(* Logix 5000 project; controller lab5BnB 5069-L306ERM rev 38.11; software revision 38.02 *)

TASK MainTask (periodic, rate 1 ms, priority 10, watchdog 1 ms) : MainProgram

MODULES
   Local : 5069-L306ERM (5069 0, rev 38.11)
       : 5069-OB16 (5069 2, rev 3.13, StandardDataDriven RPI 5 ms)
       : 5069-IB16 (5069 1, rev 2.16, StandardDataDriven RPI 5 ms)
       : vendor 1 type 115 code 320 (5069 4, rev 2.13, StandardDataDriven RPI 1 ms)
       : 5069-IF8 (5069 3, rev 3.11, StandardDataDriven RPI 1 ms)
END_MODULES

ADD_ON_INSTRUCTION Angle_Controller   (* revision 1.0 *)
VAR_INPUT
   Kp : REAL; {access None}
   Kd : REAL; {access None}
   Ki : REAL; {access None}
END_VAR
VAR_OUTPUT
   MotorInInt : REAL; {access None}
END_VAR
VAR_INPUT
   MotorVoltageInt : REAL; {access None}
   DesiredMotorAngleDeg : REAL; {access None}
END_VAR
VAR
   DERV_01 : DERIVATIVE := (Gain := 0.8, RTSTime := 1, DeltaT := 0.001);
   INTG_02 : INTEGRATOR := (IGain := 0.5, HighLimit := 4.0, LowLimit := -4.0, RTSTime := 1, Out := 1.9863874, DeltaT := 0.001);
   LPF_01 : FILTER_LOW_PASS := (WLag := 0.5, Order := 1, RTSTime := 1, DeltaT := 0.001);
   MUL_01 : FBD_MATH := (SourceA := 0.4);
   SCL_01 : SCALE := (In := 1.6115597, InRawMax := 2.8, InRawMin := -1.92, InEUMax := 90.0, InEUMin := -90.0, Limiting := 1, Out := 44.67813);
   SCL_02 : SCALE := (In := 1.9863874, InRawMax := 90.0, InRawMin := -90.0, InEUMax := -10.0, InEUMin := 10.0, Limiting := 1, Out := -0.2207098);
   SSUM_01 : SELECTED_SUMMER := (Gain1 := 1.0, Select1 := 1, Gain2 := 1.0, Select2 := 1, In3 := 1.9863874, Gain3 := 1.0, Select3 := 1, Gain4 := 1.0, Gain5 := 1.0, Gain6 := 1.0, Gain7 := 1.0, Gain8 := 1.0, Out := 1.9863874);
   SUB_01 : FBD_MATH := (SourceA := 45.0, SourceB := 45.0);
   BalanceMax : REAL := 2.8; {access None}
   BalanceMin : REAL := -1.92; {access None}
   MotorAngleDeg : REAL; {access None}
   MyError : REAL; {access None}
   PreFilter : REAL; {access None}
   PostFilter : REAL; {access None}
   __lECF02074BD2460E6 : REAL; {access None}
   __l28C6010D865A5A33 : REAL; {access None}
   __l0884565386038A91 : REAL; {access None}
   __l2DF07EE77D244EFB : REAL; {access None}
   __l1766871E0CB1B884 : REAL; {access None}
   __l0E750273472B5D8B : REAL; {access None}
   __lD887463BECBAFEBD : REAL; {access None}
   __l08A3F56F66BAD335 : REAL; {access None}
END_VAR

ROUTINE Logic   (* function block diagram *)
   SHEET 1
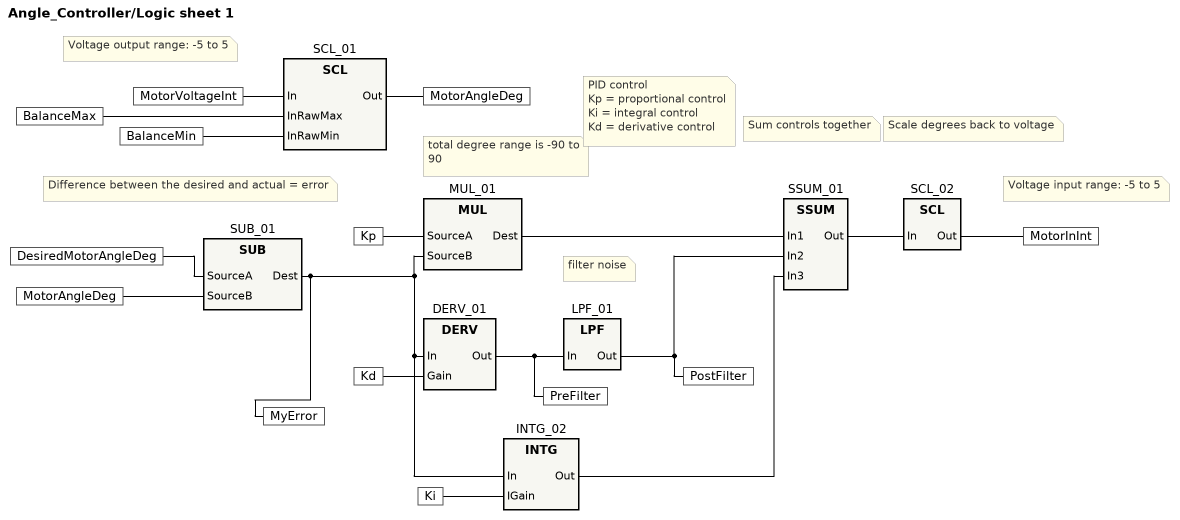
   // Difference between the desired and actual = error
   // Voltage output range: -5 to 5
   // total degree range is -90 to
   // 90
   // filter noise
   // PID control
   // Kp = proportional control
   // Ki = integral control
   // Kd = derivative control
   // Sum controls together
   // Scale degrees back to voltage
   // Voltage input range: -5 to 5
   SUB_01 : SUB(SourceA := DesiredMotorAngleDeg, SourceB := MotorAngleDeg);
   MyError := SUB_01.Dest;
   SCL_01 : SCL(In := MotorVoltageInt, InRawMax := BalanceMax, InRawMin := BalanceMin);
   MotorAngleDeg := SCL_01.Out;
   MUL_01 : MUL(SourceA := Kp, SourceB := SUB_01.Dest);
   DERV_01 : DERV(In := SUB_01.Dest, Gain := Kd);
   INTG_02 : INTG(In := SUB_01.Dest, IGain := Ki);
   PreFilter := DERV_01.Out;
   LPF_01 : LPF(In := DERV_01.Out);
   PostFilter := LPF_01.Out;
   SSUM_01 : SSUM(In1 := MUL_01.Dest, In2 := LPF_01.Out, In3 := INTG_02.Out);
   SCL_02 : SCL(In := SSUM_01.Out);
   MotorInInt := SCL_02.Out;
END_ROUTINE
END_ADD_ON_INSTRUCTION

ADD_ON_INSTRUCTION Position_Controller   (* revision 1.0 *)
VAR_INPUT
   Kp_position : REAL; {visible}
   Kd_position : REAL; {visible}
   Ki_position : REAL; {visible}
   Actual_Position : REAL; {visible}
   Desired_Position : REAL; {visible}
END_VAR
VAR_OUTPUT
   angle_out : REAL; {visible}
END_VAR
VAR
   SCL_01 : SCALE := (InRawMax := 4.5, InRawMin := -4.5, InEUMax := 7.125, InEUMin := -7.125, Limiting := 1); {access None}
   Desired_Position_Inches : DINT; {access None}
   SCL_02 : SCALE := (InRawMax := 4.5, InRawMin := -4.5, InEUMax := 7.125, InEUMin := -7.125, Limiting := 1); {access None}
   Actual_Position_Inches : DINT; {access None}
   SUB_01 : FBD_MATH := (SourceA := 45.0, SourceB := 45.0);
   MyErrorPosition : DINT; {access None}
   MUL_01 : FBD_MATH := (SourceA := 0.4);
   SCL_03 : SCALE := (In := 1.9863874, InRawMax := 7.125, InRawMin := -7.125, InEUMax := -45.0, InEUMin := 45.0, Limiting := 1, Out := -0.2207098);
   DERV_01 : DERIVATIVE := (Gain := 1.0, RTSTime := 1); {access None}
   INTG_01 : INTEGRATOR := (HighLimit := 4.0, LowLimit := -4.0, RTSTime := 1); {access None}
   SSUM_01 : SELECTED_SUMMER := (Gain1 := 1.0, Select1 := 1, Gain2 := 1.0, Select2 := 1, Gain3 := 1.0, Select3 := 1, Gain4 := 1.0, Gain5 := 1.0, Gain6 := 1.0, Gain7 := 1.0, Gain8 := 1.0); {access None}
   LPF_02 : FILTER_LOW_PASS := (WLag := 30.0, Order := 1, RTSTime := 1); {access None}
   LPF_03 : FILTER_LOW_PASS := (WLag := 30.0, Order := 1, RTSTime := 1); {access None}
   __l331A2C5B709CA8A7 : REAL; {access None}
   __l8C615611B29A5C42 : REAL; {access None}
   __l35E6236049371C91 : REAL; {access None}
   __l45EB0282393F6911 : REAL; {access None}
   __l367F46D6FCA640C7 : REAL; {access None}
END_VAR

ROUTINE Logic   (* function block diagram *)
   SHEET 1
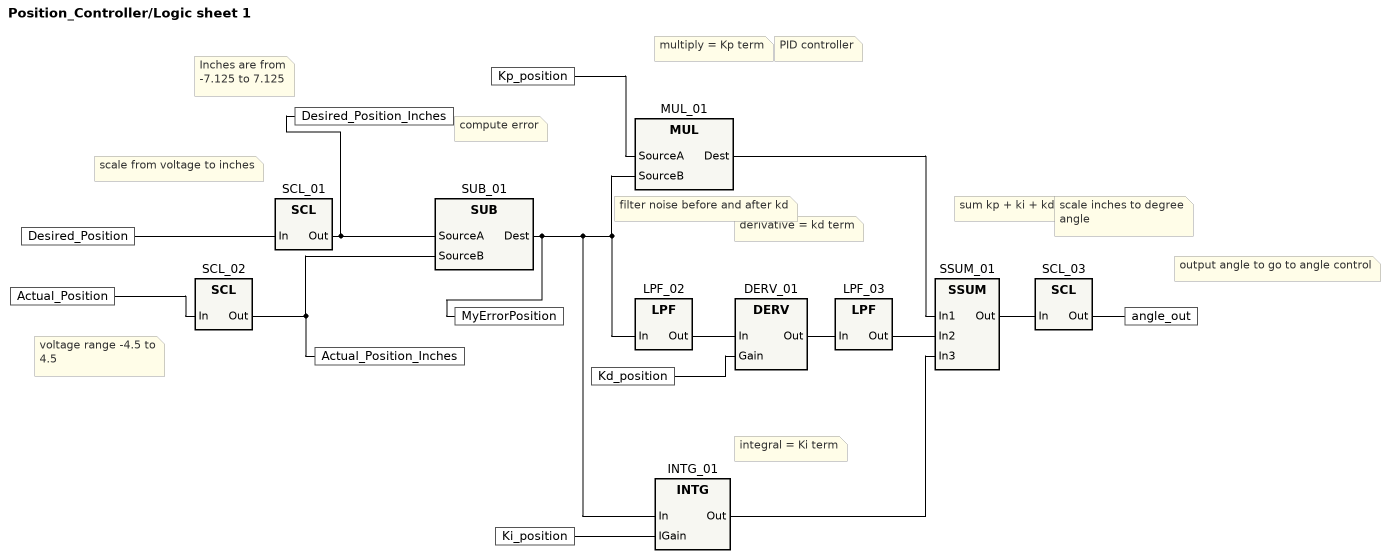
   // Inches are from
   // -7.125 to 7.125
   // voltage range -4.5 to
   // 4.5
   // scale from voltage to inches
   // compute error
   // multiply = Kp term
   // PID controller
   // integral = Ki term
   // derivative = kd term
   // filter noise before and after kd
   // sum kp + ki + kd
   // scale inches to degree
   // angle
   // output angle to go to angle control
   SCL_02 : SCL(In := Actual_Position);
   SCL_01 : SCL(In := Desired_Position);
   Desired_Position_Inches := SCL_01.Out;
   Actual_Position_Inches := SCL_02.Out;
   SUB_01 : SUB(SourceA := SCL_01.Out, SourceB := SCL_02.Out);
   MyErrorPosition := SUB_01.Dest;
   MUL_01 : MUL(SourceA := Kp_position, SourceB := SUB_01.Dest);
   LPF_02 : LPF(In := SUB_01.Dest);
   INTG_01 : INTG(In := SUB_01.Dest, IGain := Ki_position);
   DERV_01 : DERV(In := LPF_02.Out, Gain := Kd_position);
   LPF_03 : LPF(In := DERV_01.Out);
   SSUM_01 : SSUM(In1 := MUL_01.Dest, In2 := LPF_03.Out, In3 := INTG_01.Out);
   SCL_03 : SCL(In := SSUM_01.Out);
   angle_out := SCL_03.Out;
END_ROUTINE
END_ADD_ON_INSTRUCTION

VAR_GLOBAL   (* controller tags *)
   DesiredMotorAngleDeg : REAL := 6.215626;
   DesiredPosition : ALIAS FOR Local:3:I.Ch02.Data;
   DesiredPositionInches : REAL := -5.630807;
   Kd : REAL := 0.8;
   Kd_Position : REAL := 8.0;
   Ki : REAL := 0.5;
   Ki_Position : REAL := 14.0;
   Kp : REAL := 0.4;
   Kp_Position : REAL := 11.5;
   MotorAngleDeg : REAL := 4.1968155;
   MotorInInt : ALIAS FOR Local:4:O.Ch00.Data;
   MotorVoltageInt : ALIAS FOR Local:3:I.Ch00.Data;
   Position : ALIAS FOR Local:3:I.Ch01.Data;
   PositionInches : REAL := -5.626972;
END_VAR

PROGRAM MainProgram   (* main routine main *)
VAR
   Angle_Controller_01 : Angle_Controller := (Kp := 0.4, Kd := 0.8, Ki := 0.5, MotorInInt := -0.53610706, MotorVoltageInt := 0.54952836, DesiredMotorAngleDeg := 6.1429596);
   Position_Controller_01 : Position_Controller := (Kp_position := 12.0, Kd_position := 10.0, Ki_position := 10.0, Actual_Position := -3.5544348, Desired_Position := -3.5563037, angle_out := 6.1354904);
   SCL_01 : SCALE := (In := 0.5502089, InRawMax := 2.8, InRawMin := -1.92, InEUMax := 90.0, InEUMin := -90.0, Limiting := 1, Out := 4.202881);
   SCL_02 : SCALE := (In := -3.5545301, InRawMax := 4.5, InRawMin := -4.5, InEUMax := 7.125, InEUMin := -7.125, Limiting := 1, Out := -5.628006); {access None}
   SCL_03 : SCALE := (In := -3.5562074, InRawMax := 4.5, InRawMin := -4.5, InEUMax := 7.125, InEUMin := -7.125, Limiting := 1, Out := -5.630662); {access None}
END_VAR

ROUTINE main   (* function block diagram *)
   SHEET 1
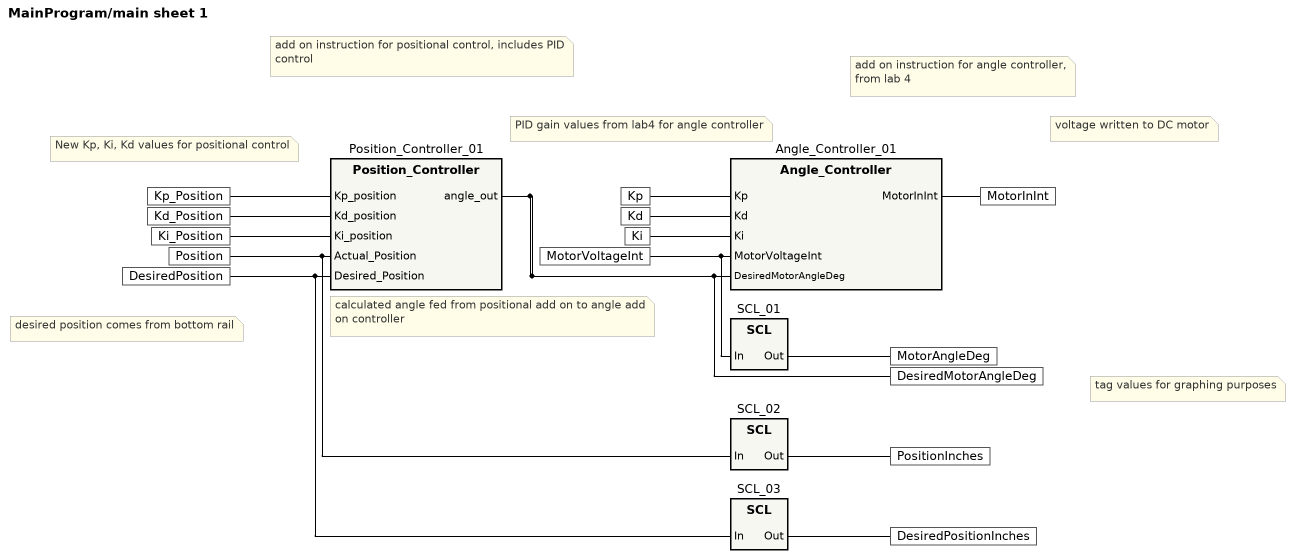
   // New Kp, Ki, Kd values for positional control
   // desired position comes from bottom rail
   // add on instruction for positional control, includes PID control
   // add on instruction for angle controller,
   // from lab 4
   // PID gain values from lab4 for angle controller
   // voltage written to DC motor
   // calculated angle fed from positional add on to angle add on controller
   // tag values for graphing purposes
   Position_Controller_01 : Position_Controller(Kp_position := Kp_Position, Kd_position := Kd_Position, Ki_position := Ki_Position, Actual_Position := Position, Desired_Position := DesiredPosition);
   Angle_Controller_01 : Angle_Controller(Kp := Kp, Kd := Kd, Ki := Ki, MotorVoltageInt := MotorVoltageInt, DesiredMotorAngleDeg := Position_Controller_01.angle_out);
   SCL_01 : SCL(In := MotorVoltageInt);
   SCL_02 : SCL(In := Position);
   SCL_03 : SCL(In := DesiredPosition);
   MotorAngleDeg := SCL_01.Out;
   DesiredMotorAngleDeg := Position_Controller_01.angle_out;
   PositionInches := SCL_02.Out;
   DesiredPositionInches := SCL_03.Out;
   MotorInInt := Angle_Controller_01.MotorInInt;
END_ROUTINE
END_PROGRAM
